SUBAPPLICATION Uebung_OPC_L19_AX (* Lokal 2x lesen: Input_I1 schreibt per PUBLISH, Output_Q1 und Output_Q2 lesen denselben Knoten (braucht FORTE mit 4diac-forte#1082) *)
  (* Standard: 61499-2; Description: Copyright (c) 2026 Meisterschulen am Ostbahnhof This program and the accompanying materials are made available under the terms of the Eclipse Public License 2.0 which is available at https://www.eclipse.org/legal/epl-2.0/ SPDX-License-Identifier: EPL-2.0 *)
  (* Version 1.0, 2026-10-18, Franz Höpfinger, Meisterschulen am Ostbahnhof, OPC-UA lokal auf einem Geraet (Meins/OPC_UA_Lokal) *)
  PACKAGE Meins::OPC_UA_Lokal;
  IMPORT Meins::OPC_UA_Lokal::const::OpcUaLokal::L19_Q_WRITE;
  IMPORT Meins::OPC_UA_Lokal::const::OpcUaLokal::L19_Q_READ;
  IMPORT logiBUS::io::DI::logiBUS_DI::Input_I1;
  IMPORT logiBUS::io::DQ::logiBUS_DO::Output_Q1;
  IMPORT logiBUS::io::DQ::logiBUS_DO::Output_Q2;
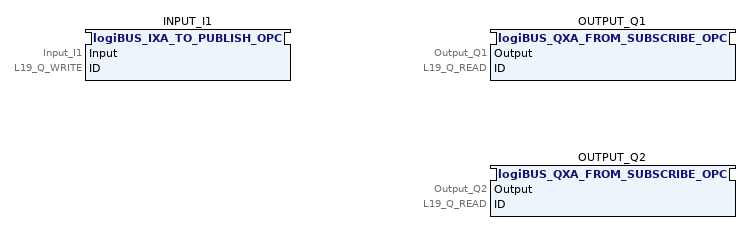
  SUBAPPS
    INPUT_I1 : MyLib::sys::logiBUS_IXA_TO_PUBLISH_OPC(Input := Input_I1, ID := L19_Q_WRITE);
    OUTPUT_Q1 : MyLib::sys::logiBUS_QXA_FROM_SUBSCRIBE_OPC(Output := Output_Q1, ID := L19_Q_READ);
    OUTPUT_Q2 : MyLib::sys::logiBUS_QXA_FROM_SUBSCRIBE_OPC(Output := Output_Q2, ID := L19_Q_READ);
  END_SUBAPPS
END_SUBAPPLICATION
